(* PLC project Untitled1, Beckhoff Automation GmbH TwinCAT PLC Control 3.5.13.21 *)
(* stored: creationDateTime 2022-12-21T13:57:08.9296352, modificationDateTime 2022-12-21T13:57:08.9336353 *)

PROGRAM MAIN
VAR
	dirM1 : BYTE := 1;
	speedM1 : WORD ;
	{attribute 'TcLinkTo' := 'TIID^Device 2 (EtherCAT)^Box 1 (sample_app)^Outputs process data mapping^Trigger'}
	dummyDataM1 AT %Q*: DWORD ;
	
	dirM2 : BYTE := 1;
	speedM2 : WORD ;
	{attribute 'TcLinkTo' := 'TIID^Device 2 (EtherCAT)^Box 2 (sample_app)^Outputs process data mapping^Trigger'}
	dummyDataM2 AT %Q*: DWORD ;
END_VAR

            dummyDataM1 := SHL(dirM1,2*8) OR speedM1 ;
dummyDataM2 := SHL(dirM2,2*8) OR speedM2 ;
          
END_PROGRAM
